// TIA Portal project "synthese" (V18)

(* hardware
DEVICE "S7-1200 station_1"  S7-1200 Station
   slot 0: "Rack_0"  S7-1200 Rack  Rack  V1.0
   slot 1: "PLC_1"  CPU 1215C DC/DC/DC  6ES7 215-1AG40-0XB0  V4.6
   slot 2: "SM 1278_1"  4SI IO link  6ES7 278-4BD32-0XB0  V2.1
   slot 3: "DI 2/DQ 2x24VDC_1"  DI2/DQ2 signal board  6ES7 223-0BD30-0XB0  V1.0
DEVICE "GSD device_1"  GSD.Device.PN
   slot 0: "Rack"  Rack  V1.0
   slot 0: "ur3ln"  V1.0  00000
      slot 0: "V1.0"  V1.0
      slot 1: "Interface"  Interface
         slot 1: "RJ45 10/100 MBit/s"  RJ45 10/100 MBit/s
   slot 5: "5_T2O General Purpose Bit Registers_1"  5_T2O General Purpose Bit Registers  1.0
      slot 0: "5_T2O General Purpose Bit Registers"  5_T2O General Purpose Bit Registers
   slot 9: "9_O2T General Purpose Registers 1_1"  9_O2T General Purpose Registers 1  1.0
      slot 0: "9_O2T General Purpose Registers 1"  9_O2T General Purpose Registers 1
DEVICE "GSD device_2"  GSD.Device.PN
   slot 0: "Rack"  Rack  V1.0
   slot 0: "vos"  default module, no PDEV  VOSxxxx-F22x  V1.8
      slot 0: "default module, no PDEV"  default module, no PDEV
      slot 1: "input module 254 byte_1"  input module 254 byte
         slot 0: "input module 254 byte"  input module 254 byte
      slot 1: "Interface"  Interface
         slot 1: "Port 1"  Port 1
      slot 2: "output module 254 byte_1"  output module 254 byte
         slot 0: "output module 254 byte"  output module 254 byte
*)

// ===== PLC "PLC_1"  CPU 1215C DC/DC/DC =====

VAR_GLOBAL   // PLC tag table "Default tag table"
   "capt 1" AT %I1.3 : Bool;
   "X5" AT %I4.0 : Bool;
   "capt 2" AT %I0.0 : Bool;
   "capt 3" AT %I1.4 : Bool;
   "X6" AT %I4.1 : Bool;
   "ind.camera 2" AT %I0.3 : Bool;
   "cobot finished" AT %I40.0 : Bool;
   "Km 1" AT %Q1.0 : Bool;
   "Led" AT %Q0.0 : Bool;
   "ind.camera 1" AT %Q0.1 : Bool;
   "cobot valid" AT %Q68.0 : Bool;
   "cobot invalid" AT %Q68.1 : Bool;
   "Led red JN" AT %Q1.5 : Bool;
   "Led yellow JN" AT %Q1.6 : Bool;
   "Led Green JN" AT %Q1.7 : Bool;
   "etat ind camera" AT %M100.0 : Bool;
   "etat finished cobot" AT %M100.1 : Bool;
   "Tag_15" AT %M10.0 : Bool;
   "Tag_16" AT %M10.1 : Bool;
   "Tag_17" AT %M10.2 : Bool;
END_VAR

// folder: System blocks/Program resources

DATA_BLOCK "IEC_Timer_0_DB"   // DB1
{ S7_Optimized_Access := 'TRUE' }
AUTHOR : Simatic
FAMILY : IEC
NAME : IEC_TMR
VERSION : 1.0
// stored: InstanceOfName IEC_TIMER
"IEC_TIMER"
BEGIN
END_DATA_BLOCK

// folder: (top level)

ORGANIZATION_BLOCK "Main"   // OB1, LAD, ProgramCycle
{ S7_Optimized_Access := 'TRUE' }
VERSION : 0.1
   VAR_INPUT
      Initial_Call : Bool;
      Remanence : Bool;
   END_VAR
BEGIN

REGION Network 1
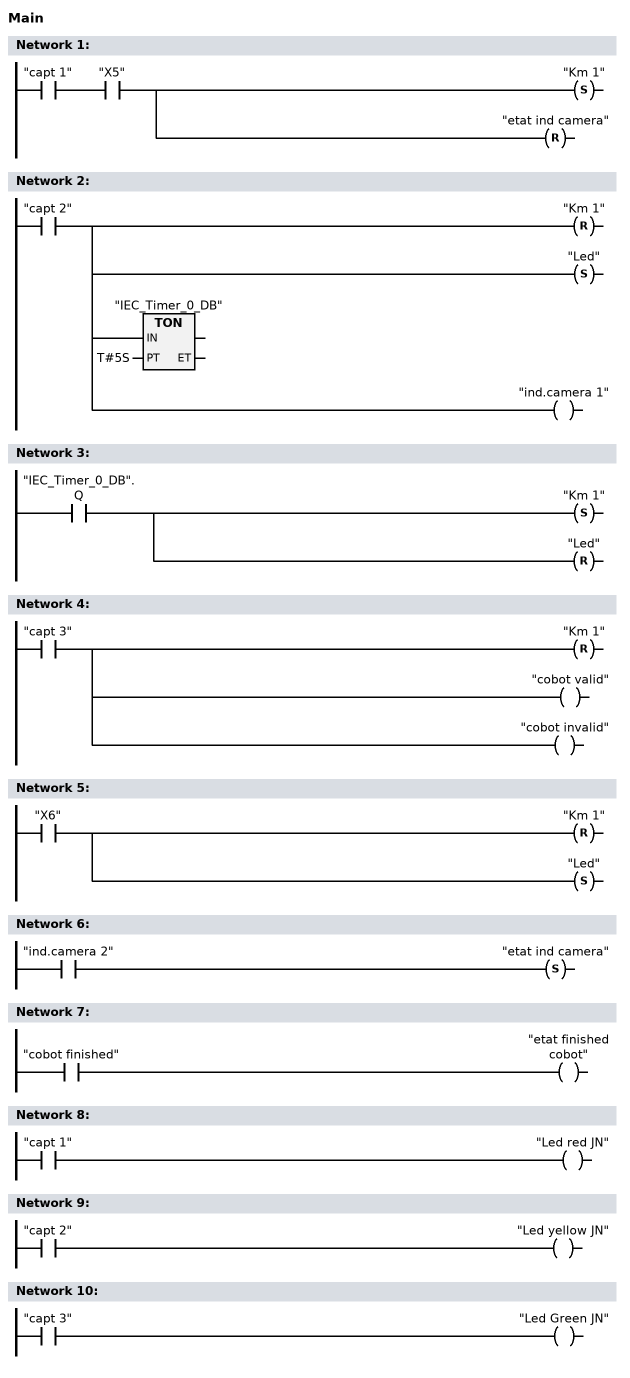
   RUNG wire#powerrail
      Contact( "capt 1" )
      Contact( "X5" )
      wire#w1
      S_Coil( "Km 1" )
   END_RUNG
   RUNG wire#w1
      R_Coil( "etat ind camera" )
   END_RUNG
   // the same network as SCL:
   IF "capt 1" AND "X5" THEN
       "Km 1" := TRUE;
       "etat ind camera" := FALSE;
   END_IF;
END_REGION

REGION Network 2
   IF "capt 2" THEN
       "Km 1" := FALSE;
       "Led" := TRUE;
   END_IF;
   "IEC_Timer_0_DB".TON(IN := "capt 2", PT := T#5S);
   "ind.camera 1" := "capt 2";
END_REGION

REGION Network 3
   RUNG wire#powerrail
      Contact( "IEC_Timer_0_DB".Q )
      wire#w1
      S_Coil( "Km 1" )
   END_RUNG
   RUNG wire#w1
      R_Coil( "Led" )
   END_RUNG
   // the same network as SCL:
   IF "IEC_Timer_0_DB".Q THEN
       "Km 1" := TRUE;
       "Led" := FALSE;
   END_IF;
END_REGION

REGION Network 4
   RUNG wire#powerrail
      Contact( "capt 3" )
      wire#w1
      R_Coil( "Km 1" )
   END_RUNG
   RUNG wire#w1
      Coil( "cobot valid" )
   END_RUNG
   RUNG wire#w1
      Coil( "cobot invalid" )
   END_RUNG
   // the same network as SCL:
   IF "capt 3" THEN "Km 1" := FALSE; END_IF;
   "cobot valid" := "capt 3";
   "cobot invalid" := "capt 3";
END_REGION

REGION Network 5
   RUNG wire#powerrail
      Contact( "X6" )
      wire#w1
      R_Coil( "Km 1" )
   END_RUNG
   RUNG wire#w1
      S_Coil( "Led" )
   END_RUNG
   // the same network as SCL:
   IF "X6" THEN
       "Km 1" := FALSE;
       "Led" := TRUE;
   END_IF;
END_REGION

REGION Network 6
   RUNG wire#powerrail
      Contact( "ind.camera 2" )
      S_Coil( "etat ind camera" )
   END_RUNG
   // the same network as SCL:
   IF "ind.camera 2" THEN "etat ind camera" := TRUE; END_IF;
END_REGION

REGION Network 7
   RUNG wire#powerrail
      Contact( "cobot finished" )
      Coil( "etat finished cobot" )
   END_RUNG
   // the same network as SCL:
   "etat finished cobot" := "cobot finished";
END_REGION

REGION Network 8
   RUNG wire#powerrail
      Contact( "capt 1" )
      Coil( "Led red JN" )
   END_RUNG
   // the same network as SCL:
   "Led red JN" := "capt 1";
END_REGION

REGION Network 9
   RUNG wire#powerrail
      Contact( "capt 2" )
      Coil( "Led yellow JN" )
   END_RUNG
   // the same network as SCL:
   "Led yellow JN" := "capt 2";
END_REGION

REGION Network 10
   RUNG wire#powerrail
      Contact( "capt 3" )
      Coil( "Led Green JN" )
   END_RUNG
   // the same network as SCL:
   "Led Green JN" := "capt 3";
END_REGION
END_ORGANIZATION_BLOCK